{attribute 'qualified_only'}
VAR_GLOBAL
    fbPmpsFileReader: FB_JsonFileToJsonDoc;
    {attribute 'pytmc' := '
        pv: @(PREFIX)DB
        io: io
    '}
    fbStandardPMPSDB: FB_Standard_PMPSDB;
END_VAR

(* stored: Version 1.1.0.1, ProductVersion 3.1.4022.18
   GVL MOTION_GVL: Id {7b3cfad1-1f36-4ed6-b576-62277c19b2b2} *)
